FUNCTION_BLOCK FB_Blikjesband IMPLEMENTS ITF_Blikjesband
VAR_INPUT
END_VAR
VAR_OUTPUT
END_VAR
VAR
END_VAR

{warning 'Add method implementation '}
METHOD Aborted : BOOL
END_METHOD

{warning 'Add method implementation '}
METHOD Aborting : BOOL
END_METHOD

{warning 'Add method implementation '}
METHOD Clearing : BOOL
END_METHOD

{warning 'Add method implementation '}
METHOD Execute : BOOL
END_METHOD

{warning 'Add method implementation '}
METHOD Held : BOOL
END_METHOD

{warning 'Add method implementation '}
METHOD Holding : BOOL
END_METHOD

{warning 'Add method implementation '}
METHOD Idle : BOOL
END_METHOD

{warning 'Add method implementation '}
METHOD Resetting : BOOL
END_METHOD

{warning 'Add method implementation '}
METHOD Starting : BOOL
END_METHOD

{warning 'Add method implementation '}
METHOD Stopped : BOOL
END_METHOD

{warning 'Add method implementation '}
METHOD Stopping : BOOL
END_METHOD

{warning 'Add method implementation '}
METHOD Suspended : BOOL
END_METHOD

{warning 'Add method implementation '}
METHOD Suspending : BOOL
END_METHOD

{warning 'Add method implementation '}
METHOD Unholding : BOOL
END_METHOD

{warning 'Add method implementation '}
METHOD Unsuspending : BOOL
END_METHOD

END_FUNCTION_BLOCK

(* stored: Version 1.1.0.1
   POU FB_Blikjesband: Id {50ab0147-870b-4937-87bd-ef941e378017}, SpecialFunc None
   Folder Methods: Id {0c50d0d5-ba27-478e-b2d5-2bc613b9db20}
   Method Aborted: Id {cf1f3de9-2227-4dc2-bc44-19c7bde3462b}
   Method Aborting: Id {e2516ec8-70d9-41d5-bbc5-0c4700635e54}
   Method Clearing: Id {39c60839-9082-445d-90ff-0e60501d4066}
   Method Execute: Id {aa06be4f-f4fc-4af0-927c-8e1ca37728fc}
   Method Held: Id {31e1809f-2cda-4718-94e8-9049b4e88853}
   Method Holding: Id {3ea68ff6-7c42-42e7-abd6-2bdc373272be}
   Method Idle: Id {615dfa91-b11b-4774-ac7a-ab8fbaf1eac6}
   Method Resetting: Id {faa8be60-8ba0-4fbf-8818-0d0c0aa443e6}
   Method Starting: Id {4219dfd1-b119-4acb-a3b5-a41aa59efcf2}
   Method Stopped: Id {84165a36-9fa6-4f5c-910b-cdf58fead66a}
   Method Stopping: Id {a5baaab6-55e7-4141-9d6b-8b12a39c69ad}
   Method Suspended: Id {d504ec83-13ae-44e8-96ef-7f958e37d3fc}
   Method Suspending: Id {5fd4895e-7660-4cb3-8d98-8fc78d8948b6}
   Method Unholding: Id {a5a70ae8-1b02-413b-9c51-a635862c2ecd}
   Method Unsuspending: Id {74f5fec4-1978-4558-b9a8-b0cda332b4be} *)
